Fanuc KAREL source: kt00048.KL

-- PROVISIONAL review KL for V1013-1; original PC SHA256 5fac9843858cc6c0a74672d89afdf6a80996552cff14631e6fea422bc16e96f7
-- Incomplete behavior may be omitted. Consult companion uncertainty JSON. Do not deploy.
PROGRAM KT00048
%NOLOCKGROUP
VAR
  R1 : REAL
  OUT : REAL
-- UNRESOLVED_DECL H2 type=002017
BEGIN
  -- UNRESOLVED_PC offsets 5-16; opcodes 2E,23
  -- UNRESOLVED_PC offsets 21-35; opcodes 2E,22,9D,33,B4
  -- UNRESOLVED_PC offsets 40-63; opcodes 21,22,9D,33,B3,64,6A,23
  -- UNRESOLVED_PC offsets 68-72; opcodes 7F
END KT00048
